// PlcTask 每 2 ms 调用；先刷新反馈，再判组条件，再轨迹，最后基础轴块。
// 每轴的 NC 引用、ADS 数据、参数及传感器索引必须一一对应。
PROGRAM MAIN
VAR
    fbAxisConfig : FB_AxisConfig; // 独立轴配置入口，仅在有效空闲时应用本块的虚拟轴参数。
    fbAxis1 : FB_AxisControl; // 轴1基础控制实例，固定对应 GVL_sy.axis[1] 和 GVL_axis.Axis1。
    fbAxis2 : FB_AxisControl; // 轴2基础控制实例，固定对应 GVL_sy.axis[2] 和 GVL_axis.Axis2。
    fbAxis3 : FB_AxisControl; // 轴3基础控制实例，固定对应 GVL_sy.axis[3] 和 GVL_axis.Axis3。
    fbAxis4 : FB_AxisControl; // 轴4基础控制实例，固定对应 GVL_sy.axis[4] 和 GVL_axis.Axis4。
    fbAuthority : FB_ControlAuthority; // 三站控制权仲裁实例，处理申请、释放、心跳和交接锁。
    aCommandGate : ARRAY[1..4] OF FB_AxisCommandGate; // 四轴手动命令门，只向对应轴转交当前持有站的有效命令。
    xControlBusy : BOOL; // 实际运动、轨迹或轴块忙的汇总，作为禁止控制权交接的判据。
    nManualStation : UINT; // 本扫描允许读取的站号；0 时命令门清除旧请求。
    fbTrajectory : FB_FourAxisTrajectory; // 四轴点位接收、拼表、校验及轨迹执行实例。
    fbHmiFeedback : FB_HmiFeedback; // 四轴执行结果发布到 switch 只读监控接口。
    xAllEnabled : BOOL; // 四轴使能反馈，用于运行中判断是否掉使能。
    xAxesReady : BOOL; // 轨迹启动就绪：四轴使能、回原、静止且不在停车。
    nAbortReason : UINT; // 本扫描首个联停原因；0 表示没有联停请求。
    xAbort : BOOL; // 整组联停请求，汇总许可丢失、撤使能、命令冲突及限位等条件。
    xAxisFault : BOOL; // 任一基础轴错误或 NC 错误、I/O 无效，供轨迹块判断故障。
    i : INT; // 四轴状态汇总的循环轴号，范围 1～4。
END_VAR

// 当前仅用于虚拟轴软件调试，明确给出运行许可。
// 接实机前必须将下一行替换为现场安全继电器的运行允许反馈。
GVL_motion.xMotionPermit := TRUE;

// 刷新四轴实际状态；只读取 NC 反馈，不要求持有控制权。
A01_ReadAxisStatus();

// 汇总交接条件并处理控制权；写入 GVL_control 仲裁反馈。
A02_ControlAuthority();

// 轴配置单独处理，使用当前运动锁和现有空闲反馈。
fbAxisConfig();

// 取出授权站手动命令；通过命令门写入 GVL_axis 命令字段。
A03_ManualCommands();

// 汇总轨迹联锁并调用原轨迹块；更新 GVL_motion 轨迹状态。
A04_TrajectoryControl();

// 调用四轴基础控制；更新 NC 控制输出及 GVL_axis 实际反馈。
A05_ManualAxes();

// 发布本扫描执行后的反馈；只写 GVL_HMI，不产生运动命令。
A06_PublishFeedback();

ACTION A01_ReadAxisStatus:
// 刷新四轴实际状态；只读取 NC 反馈，不要求持有控制权。
// 先统一刷新轴状态，再决定四轴本周期的共同轨迹帧。
FOR i := 1 TO 4 DO
 GVL_sy.axis[i].ReadStatus();
 END_FOR
END_ACTION

ACTION A02_ControlAuthority:
// 汇总交接条件并处理控制权；写入 GVL_control 仲裁反馈。
// 运行锁：点动、回原、轨迹、停止/退出及未消费的运动命令都阻止交接。
// 使用 NC 状态、实际速度和轴块 Busy；I/O 无效单独发布，不能冒充运动占用。
xControlBusy := GVL_motion.xBusy OR GVL_axis.Axis1.xBusy OR GVL_axis.Axis2.xBusy
    OR GVL_axis.Axis3.xBusy OR GVL_axis.Axis4.xBusy;
GVL_control.xFeedbackInvalid := FALSE;
FOR i := 1 TO 4 DO
    xControlBusy := xControlBusy OR GVL_sy.axis[i].Status.Moving
        OR GVL_sy.axis[i].Status.Homing OR GVL_sy.axis[i].Status.Stopping
        OR GVL_sy.axis[i].Status.ExtSetPointGenEnabled
        OR (ABS(GVL_sy.axis[i].NcToPlc.ActVelo) > 0.000001);
    GVL_control.xFeedbackInvalid := GVL_control.xFeedbackInvalid OR GVL_sy.axis[i].Status.IoDataInvalid;
END_FOR
fbAuthority(xMotionBusy := xControlBusy, xFeedbackInvalid := GVL_control.xFeedbackInvalid);
END_ACTION

ACTION A03_ManualCommands:
// 四个命令门共用本扫描的授权结果，各自读取对应轴的邮箱。
// 交接扫描仍清除旧请求，新持有者须在确认授权后重新发命令。
nManualStation := 0;
IF GVL_control.xCanCommand AND NOT GVL_control.xOwnerChanged THEN
    nManualStation := GVL_control.nOwner;
END_IF
aCommandGate[1](Data := GVL_axis.Axis1, nStation := nManualStation, nAxis := 1, xStop := GVL_control.xStopOwner);
aCommandGate[2](Data := GVL_axis.Axis2, nStation := nManualStation, nAxis := 2, xStop := GVL_control.xStopOwner);
aCommandGate[3](Data := GVL_axis.Axis3, nStation := nManualStation, nAxis := 3, xStop := GVL_control.xStopOwner);
aCommandGate[4](Data := GVL_axis.Axis4, nStation := nManualStation, nAxis := 4, xStop := GVL_control.xStopOwner);
END_ACTION

ACTION A04_TrajectoryControl:
// 汇总轨迹联锁并调用原轨迹块；更新 GVL_motion 轨迹状态。
// 基础轴块在轨迹块之后调用，此处使用上一扫描的使能反馈。
xAllEnabled := GVL_axis.Axis1.xEnabled AND GVL_axis.Axis2.xEnabled AND GVL_axis.Axis3.xEnabled AND GVL_axis.Axis4.xEnabled;
xAxisFault := GVL_axis.Axis1.xError OR GVL_axis.Axis2.xError  OR GVL_axis.Axis3.xError OR GVL_axis.Axis4.xError;
// 按许可、控制权、使能、停止、手动冲突、限位的顺序取第一个联停原因。
// 当前持有站发出的整组停止命令，由轨迹块走正常停车流程。
nAbortReason := 0;
IF NOT GVL_motion.xMotionPermit THEN nAbortReason := 1;
ELSIF NOT GVL_control.xCanCommand THEN nAbortReason := 2;
ELSIF (GVL_motion.xBusy AND NOT xAllEnabled)
    OR NOT GVL_axis.Axis1.xStart OR NOT GVL_axis.Axis2.xStart
    OR NOT GVL_axis.Axis3.xStart OR NOT GVL_axis.Axis4.xStart THEN nAbortReason := 3;
ELSIF (GVL_axis.Axis1.xStop OR GVL_axis.Axis2.xStop OR GVL_axis.Axis3.xStop OR GVL_axis.Axis4.xStop)
    AND NOT ((GVL_motion.nCommandStation = GVL_control.nOwner) AND GVL_motion.xStop) THEN nAbortReason := 4;
ELSIF GVL_axis.Axis1.jogz OR GVL_axis.Axis1.jogf OR GVL_axis.Axis1.gohome OR GVL_axis.Axis1.reset
    OR GVL_axis.Axis2.jogz OR GVL_axis.Axis2.jogf OR GVL_axis.Axis2.gohome OR GVL_axis.Axis2.reset
    OR GVL_axis.Axis3.jogz OR GVL_axis.Axis3.jogf OR GVL_axis.Axis3.gohome OR GVL_axis.Axis3.reset
    OR GVL_axis.Axis4.jogz OR GVL_axis.Axis4.jogf OR GVL_axis.Axis4.gohome OR GVL_axis.Axis4.reset THEN
    nAbortReason := 5;
END_IF
// 启动就绪才要求回原和静止，运行中用使能反馈判断掉使能。
xAxesReady := xAllEnabled;
FOR i := 1 TO 4 DO
    xAxesReady := xAxesReady AND GVL_sy.axis[i].Status.Homed AND GVL_sy.axis[i].Status.StandStill AND NOT GVL_sy.axis[i].Status.Stopping;
    xAxisFault := xAxisFault OR GVL_sy.axis[i].Status.Error OR GVL_sy.axis[i].Status.IoDataInvalid;
    IF (nAbortReason = 0) AND (GVL_motion.axPositiveLimit[i] OR GVL_motion.axNegativeLimit[i]
        OR GVL_sy.axis[i].Status.SoftLimitMinExceeded OR GVL_sy.axis[i].Status.SoftLimitMaxExceeded) THEN
        nAbortReason := 6;
    END_IF
END_FOR
xAbort := nAbortReason <> 0;
// 轨迹块先更新组状态和 xBusy，后面的基础块在本扫描就能据此禁止手动抢占。
// 全部下发后的统一拼表状态 5 不置 xBusy，不占用基础轴控制。
fbTrajectory(Axes := GVL_sy.axis, xAxesReady := xAxesReady, xAbort := xAbort, xAxisFault := xAxisFault, nAbortReason := nAbortReason);
END_ACTION

ACTION A05_ManualAxes:
// 调用四轴基础控制；更新 NC 控制输出及 GVL_axis 实际反馈。
// 四个实例各自保存 Power/Jog/Home/Stop/Reset 的状态，便于逐轴打断点。
// 四个基础实例每扫描都调用，持续更新异步 MC 块 Busy/Done/Error。
// Axis1..4 固定对应 NC 引用 [1]..[4]，不通过选中轴号复用一个实例。
fbAxis1(Axis := GVL_sy.axis[1], Data := GVL_axis.Axis1, Config := GVL_motion.aConfig[1],
    xPermit := GVL_motion.xMotionPermit AND GVL_control.xCanCommand, xPositiveLimit := GVL_motion.axPositiveLimit[1],
    xNegativeLimit := GVL_motion.axNegativeLimit[1], xHomeSensor := GVL_motion.axHomeSensor[1],
    xGroupBusy := GVL_motion.xBusy);
fbAxis2(Axis := GVL_sy.axis[2], Data := GVL_axis.Axis2, Config := GVL_motion.aConfig[2],
    xPermit := GVL_motion.xMotionPermit AND GVL_control.xCanCommand, xPositiveLimit := GVL_motion.axPositiveLimit[2],
    xNegativeLimit := GVL_motion.axNegativeLimit[2], xHomeSensor := GVL_motion.axHomeSensor[2],
    xGroupBusy := GVL_motion.xBusy);
fbAxis3(Axis := GVL_sy.axis[3], Data := GVL_axis.Axis3, Config := GVL_motion.aConfig[3],
    xPermit := GVL_motion.xMotionPermit AND GVL_control.xCanCommand, xPositiveLimit := GVL_motion.axPositiveLimit[3],
    xNegativeLimit := GVL_motion.axNegativeLimit[3], xHomeSensor := GVL_motion.axHomeSensor[3],
    xGroupBusy := GVL_motion.xBusy);
fbAxis4(Axis := GVL_sy.axis[4], Data := GVL_axis.Axis4, Config := GVL_motion.aConfig[4],
    xPermit := GVL_motion.xMotionPermit AND GVL_control.xCanCommand, xPositiveLimit := GVL_motion.axPositiveLimit[4],
    xNegativeLimit := GVL_motion.axNegativeLimit[4], xHomeSensor := GVL_motion.axHomeSensor[4],
    xGroupBusy := GVL_motion.xBusy);
END_ACTION

ACTION A06_PublishFeedback:
// 发布本扫描执行后的反馈；只写 GVL_HMI，不产生运动命令。
// 所有基础块本周期输出更新后，再发布 HMI 状态；避免把请求位误当成执行反馈。
fbHmiFeedback();
END_ACTION

END_PROGRAM

(* stored: Version 1.1.0.1
   POU MAIN: Id {df6a7805-2d1f-401a-b50b-7126627d78b7}, SpecialFunc None
   Action A01_ReadAxisStatus: Id {d342207c-f231-5ee1-99f1-05ad1db0ec87}
   Action A02_ControlAuthority: Id {3eeb1f59-5728-51cf-b201-23836cbf5d99}
   Action A03_ManualCommands: Id {455d291c-6bbf-5830-8f93-78839db9156a}
   Action A04_TrajectoryControl: Id {1d20d96a-49bd-5fb3-9b5c-92dd45de2540}
   Action A05_ManualAxes: Id {e283efde-06ca-5b80-bffe-6ba54f46393f}
   Action A06_PublishFeedback: Id {1ee1214a-0779-5158-9078-6f391e452af9} *)
